Fanuc KAREL source: kc00041.KL

-- PROVISIONAL review KL for V770-1; original PC SHA256 4a75ddb66af0bb3a1b8ba5b0396bc6df869e47ba5e79e879aa93335f3083948b
-- Incomplete behavior may be omitted. Consult companion uncertainty JSON. Do not deploy.
PROGRAM KC00041
%NOLOCKGROUP
BEGIN
  -- UNRESOLVED_PC offsets 5-33; opcodes 27,22,22,22,22,31
  -- UNRESOLVED_PC offsets 38-42; opcodes 7F
END KC00041
